Fanuc KAREL source: kd00022.KL

-- PROVISIONAL review KL for V1013-1; original PC SHA256 7b83e7b8f417eb635d9ef1a48d5c14f71e8f6bb26466e07f7661abea11e99437
-- Incomplete behavior may be omitted. Consult companion uncertainty JSON. Do not deploy.
PROGRAM KD00022
%NOLOCKGROUP
VAR
  I : INTEGER
  J : INTEGER
  B : BOOLEAN
  R : REAL
  S : STRING[80]
-- UNRESOLVED_DECL SAVED type=fd0010
BEGIN
  -- UNRESOLVED_PC offsets 5-12; opcodes 9D,23
  -- UNRESOLVED_PC offsets 17-21; opcodes 7F
END KD00022
